(* IEC 61131-3 sources: plc-process-lib/src/DUTs/Motor, 6 files *)

(* ---- E_MotorAlarm.dut.st ---- *)
// Назначение: индексы слотов тревог двигателя; слоты 6–7 — только у FB_MotorVfd.
//             Нестрогое перечисление: им индексируются массивы.
// Автор:      kr0nsch
// Версия:     0.1.0
// Документ:   docs/fb/FB_Motor.md
{attribute 'qualified_only'}
TYPE E_MotorAlarm :
(
    FailToStart    := 0,   // нет ОС за tFbStart
    FeedbackLost   := 1,   // ОС пропала в работе
    FailToStop     := 2,   // ОС не пропала за tFbStop
    UncommandedRun := 3,   // ОС без команды
    ExtFault       := 4,   // внешняя авария
    InterlockTrip  := 5,   // останов блокировкой в работе
    CommLoss       := 6,   // потеря связи с ПЧ
    SpeedDeviation := 7    // рассогласование задания и фактической скорости ПЧ
) UINT;
END_TYPE

(* ---- E_MotorState.dut.st ---- *)
// Назначение: состояние двигателя (FB_Motor, FB_MotorVfd).
// Автор:      kr0nsch
// Версия:     0.1.0
// Документ:   docs/fb/FB_Motor.md
{attribute 'qualified_only'}
{attribute 'strict'}
TYPE E_MotorState :
(
    Stopped  := 0,
    Starting := 1,   // команда подана, ждём ОС
    Running  := 2,
    Stopping := 3,   // команда снята, ждём пропадания ОС
    Fault    := 4    // отказ: выходы сняты, ждём Reset (или восстановления связи с ПЧ)
) INT;
END_TYPE

(* ---- ST_MotorCfg.dut.st ---- *)
// Назначение: параметры двигателя (FB_Motor и FB_MotorVfd; Persistent Variables приложения,
//             VAR_IN_OUT CONSTANT stCfg). Значения по умолчанию проходят CheckConfig. Маски
//             по умолчанию 16#FFFF: забытая маска даёт «блокирует», а не «молча игнорирует».
//             Тип лежит в Persistent Variables приложения и заморожен в пределах 1.x (A-13).
// Автор:      kr0nsch
// Версия:     0.1.0
// Документ:   docs/fb/FB_Motor.md
{attribute 'qualified_only'}
TYPE ST_MotorCfg :
STRUCT
    xFbUsed            : BOOL := TRUE;      // ОС «в работе» подключена
    tFbStart           : TIME := T#5S;      // ожидание ОС при пуске (для УПП — не меньше времени разгона)
    tFbStop            : TIME := T#5S;      // ожидание пропадания ОС при останове (выбег)
    tFbLossFilter      : TIME := T#500MS;   // фильтр пропадания ОС в работе
    tExtFaultFilter    : TIME := T#200MS;   // фильтр внешней аварии
    tMinRun            : TIME := T#0S;      // мин. время работы — только для остановов от автоматики
    tMinStop           : TIME := T#0S;      // мин. пауза перед пуском (также после старта ПЛК и провала питания)
    uiMaxStartsPerHour : UINT := 0;         // 0 — без ограничения; не больше STARTS_WINDOW_MAX
    tResetWindow       : TIME := T#3S;      // окно снятия причин после Reset (сброс УПП/ПЧ)
    tResetPulse        : TIME := T#1S;      // длительность импульса xQReset; не больше tResetWindow
    wInterlockMask     : WORD := 16#FFFF;   // какие биты wInterlock действуют
    wPermitMask        : WORD := 16#FFFF;   // какие биты wPermit обязательны для пуска
    udiMaintInterval_h : UDINT := 0;        // ТО по наработке, ч; 0 — нет
    udiMaintStarts     : UDINT := 0;        // ТО по числу пусков; 0 — нет
    stVfd              : ST_VfdCfg;         // только FB_MotorVfd
    udiAlarmIdBase     : UDINT := 0;        // номер первой тревоги устройства (dev_no * 10)
    astAlarm           : ARRAY[0..GVL_Const.DEV_ALARMS_MAX - 1] OF ST_AlarmCfg := [
        (ePriority := E_AlarmPriority.Medium),    // 0 FailToStart
        (ePriority := E_AlarmPriority.Medium),    // 1 FeedbackLost
        (ePriority := E_AlarmPriority.High),      // 2 FailToStop — механизм не остановить из ПЛК
        (ePriority := E_AlarmPriority.High),      // 3 UncommandedRun
        (ePriority := E_AlarmPriority.Medium),    // 4 ExtFault
        (ePriority := E_AlarmPriority.None),      // 5 InterlockTrip — у причины обычно своя тревога
        (ePriority := E_AlarmPriority.Medium),    // 6 CommLoss (ПЧ)
        (ePriority := E_AlarmPriority.Low)];      // 7 SpeedDeviation (ПЧ)
END_STRUCT
END_TYPE

(* ---- ST_MotorCmd.dut.st ---- *)
// Назначение: команды HMI/SCADA двигателя (FB_Motor и FB_MotorVfd, VAR_IN_OUT stCmd).
// Автор:      kr0nsch
// Версия:     0.1.0
// Документ:   docs/fb/FB_Motor.md
{attribute 'qualified_only'}
TYPE ST_MotorCmd :
STRUCT
    stCommon     : ST_DeviceCmd;
    xStart       : BOOL;   // импульс: пуск (Manual; в Auto — RejectedMode)
    xStop        : BOOL;   // импульс: стоп (в Auto — переход в Manual и стоп)
    xResetMaint  : BOOL;   // импульс: обнулить счётчики «с последнего ТО»
    rSpeedSp_pct : REAL;   // ПЧ: задание скорости в Manual, %; в Auto/Local/OOS ФБ пишет сюда текущее
END_STRUCT
END_TYPE

(* ---- ST_MotorSts.dut.st ---- *)
// Назначение: состояние двигателя для HMI/SCADA (и для FB_MotorVfd). 68 байт, 34 регистра
//             Modbus: только 16- и 32-битные поля без скрытого выравнивания.
// Автор:      kr0nsch
// Версия:     0.1.0
// Документ:   docs/fb/FB_Motor.md
{attribute 'qualified_only'}
TYPE ST_MotorSts :
STRUCT
    stCommon          : ST_DeviceSts;   // 0..27; eDevType = MotorVfd — фейсплейт показывает блок ПЧ
    eState            : E_MotorState;   // 28
    wInterlock        : WORD;    // 30: действующие блокировки (wInterlock AND wInterlockMask)
    wPermitMissing    : WORD;    // 32: недостающие разрешения (wPermitMask AND NOT wPermit)
    uiFirstOut        : UINT;    // 34: номер бита первой сработавшей блокировки 0..15; NO_FIRST_OUT — нет
    uiInhibitRemain_s : UINT;    // 36: до снятия запрета пуска (пауза, лимит пусков), с, вверх, <= UINT_MAX
    uiStartsLastHour  : UINT;    // 38: пусков за скользящий час
    rRunTime_h        : REAL;    // 40: наработка всего, ч
    udiStarts         : UDINT;   // 44: пусков всего
    rRunTimeMaint_h   : REAL;    // 48: наработка с последнего ТО, ч
    udiStartsMaint    : UDINT;   // 52: пусков с последнего ТО
    rSpeedRef_pct     : REAL;    // 56: задание на ПЧ после ограничений и рампы, % (0 у прямого пуска)
    rSpeedAct_pct     : REAL;    // 60: фактическая скорость, % (0 у прямого пуска)
    udiRunCurrent_s   : UDINT;   // 64: текущая непрерывная работа, с; 0, пока стоит
END_STRUCT
END_TYPE

(* ---- ST_VfdCfg.dut.st ---- *)
// Назначение: параметры преобразователя частоты (поле stVfd в ST_MotorCfg); используется
//             только FB_MotorVfd.
//             Тип лежит в Persistent Variables приложения и заморожен в пределах 1.x (A-13).
// Автор:      kr0nsch
// Версия:     0.1.0
// Документ:   docs/fb/FB_MotorVfd.md
{attribute 'qualified_only'}
TYPE ST_VfdCfg :
STRUCT
    rSpeedMin_pct    : REAL := 0.0;    // мин. задание в работе, % (по данным насоса и двигателя)
    rSpeedMax_pct    : REAL := 100.0;  // макс. задание, %
    rRampUp_pctps    : REAL := 0.0;    // ограничение роста задания, %/с; 0 — нет (работают рампы ПЧ)
    rRampDown_pctps  : REAL := 0.0;    // ограничение спада задания, %/с; 0 — нет
    xFbFromComm      : BOOL := TRUE;   // ОС «в работе» — из слова состояния ПЧ (xVfdRunning); FALSE — DI xFbRun
    xCommLossIsFault : BOOL := TRUE;   // FALSE — пуск/стоп заведены проводами, по Modbus только задание
    tCommLoss        : TIME := T#3S;   // фильтр потери связи
    rSpeedDev_pct    : REAL := 10.0;   // допустимое рассогласование задание/факт; 0 — контроль выключен
    tSpeedDev        : TIME := T#10S;  // задержка рассогласования
END_STRUCT
END_TYPE
